(* IEC 61131-3 sources: llm-plc-st-eval/data/processed_definitivo/gpt-4o-2024-08-06/I8/zero_shot, 3 files *)

(* ---- ejec_1.st ---- *)
FUNCTION_BLOCK FB_Compresor
VAR_INPUT
    pOilOk : BOOL;        // Presión de aceite correcta
    tempOk : BOOL;        // Temperatura correcta
    sinAlm : BOOL;        // Sin alarmas
    btnMarcha : BOOL;     // Botón de marcha
    btnParo : BOOL;       // Botón de paro
END_VAR

VAR_OUTPUT
    comp : BOOL;          // Salida del compresor
    causaBloqueo : INT;   // Causa del bloqueo
END_VAR

VAR
    pOilOkTimer : TON;    // Temporizador para presión de aceite
    btnMarchaPrev : BOOL; // Estado previo del botón de marcha
END_VAR

// Inicialización del temporizador
pOilOkTimer(IN := pOilOk, PT := T#3S);

// Evaluación de los permisivos
IF NOT pOilOkTimer.Q THEN
    causaBloqueo := 1; // Falta presión de aceite
ELSIF NOT tempOk THEN
    causaBloqueo := 2; // Falta temperatura correcta
ELSIF NOT sinAlm THEN
    causaBloqueo := 3; // Alarma activa
ELSE
    causaBloqueo := 0; // Todos los permisivos están bien
END_IF

// Lógica de control del compresor
IF btnParo THEN
    comp := FALSE; // Parar el compresor
ELSIF NOT comp THEN
    // Arrancar el compresor solo si se presiona btnMarcha y todos los permisivos están bien
    IF btnMarcha AND NOT btnMarchaPrev AND causaBloqueo = 0 THEN
        comp := TRUE;
    END_IF
END_IF

// Actualizar el estado previo del botón de marcha
btnMarchaPrev := btnMarcha;
END_FUNCTION_BLOCK

(* ---- ejec_2.st ---- *)
FUNCTION_BLOCK FB_Compresor
VAR_INPUT
    pOilOk : BOOL;       // Presión de aceite correcta
    tempOk : BOOL;       // Temperatura correcta
    sinAlm : BOOL;       // Ausencia de alarmas
    btnMarcha : BOOL;    // Botón de marcha
    btnParo : BOOL;      // Botón de paro
END_VAR

VAR_OUTPUT
    comp : BOOL;         // Estado del compresor
    causaBloqueo : INT;  // Causa de bloqueo
END_VAR

VAR
    pOilOkTimer : TON;   // Temporizador para presión de aceite
    marchaPrev : BOOL;   // Estado anterior de btnMarcha
END_VAR

// Inicialización del temporizador
pOilOkTimer(IN := pOilOk, PT := T#3S);

// Lógica para determinar la causa de bloqueo
IF NOT pOilOk THEN
    causaBloqueo := 1; // Falta presión de aceite
ELSIF NOT tempOk THEN
    causaBloqueo := 2; // Falta temperatura correcta
ELSIF NOT sinAlm THEN
    causaBloqueo := 3; // Hay alarmas activas
ELSE
    causaBloqueo := 0; // No hay bloqueos
END_IF;

// Lógica de control del compresor
IF btnParo THEN
    comp := FALSE; // Parar el compresor si se pulsa btnParo
ELSIF comp THEN
    // Mantener el compresor en marcha si está en marcha y no hay bloqueos
    IF NOT (pOilOkTimer.Q AND tempOk AND sinAlm) THEN
        comp := FALSE; // Parar si se pierde algún permisivo
    END_IF;
ELSE
    // Arrancar el compresor si se pulsa btnMarcha y se cumplen los permisivos
    IF btnMarcha AND NOT marchaPrev AND pOilOkTimer.Q AND tempOk AND sinAlm THEN
        comp := TRUE;
    END_IF;
END_IF;

// Actualizar el estado anterior de btnMarcha
marchaPrev := btnMarcha;

END_FUNCTION_BLOCK

(* ---- ejec_3.st ---- *)
FUNCTION_BLOCK FB_Compresor
VAR
    // Entradas
    pOilOk : BOOL;       // Presión de aceite correcta
    tempOk : BOOL;       // Temperatura correcta
    sinAlm : BOOL;       // Sin alarmas
    btnMarcha : BOOL;    // Botón de marcha
    btnParo : BOOL;      // Botón de paro

    // Salidas
    comp : BOOL;         // Estado del compresor
    causaBloqueo : INT;  // Causa de bloqueo

    // Variables internas
    pOilOkTimer : TON;   // Temporizador para presión de aceite
    marchaLatch : BOOL;  // Latch para mantener el compresor en marcha
END_VAR

// Inicialización del temporizador
pOilOkTimer(IN := pOilOk, PT := T#3S);

// Lógica de causa de bloqueo
IF NOT pOilOkTimer.Q THEN
    causaBloqueo := 1; // Falta presión de aceite
ELSIF NOT tempOk THEN
    causaBloqueo := 2; // Falta temperatura correcta
ELSIF NOT sinAlm THEN
    causaBloqueo := 3; // Hay alarmas activas
ELSE
    causaBloqueo := 0; // No hay bloqueos
END_IF;

// Lógica de arranque y paro del compresor
IF btnParo THEN
    marchaLatch := FALSE; // Parar el compresor
ELSIF btnMarcha AND NOT marchaLatch AND (causaBloqueo = 0) THEN
    marchaLatch := TRUE; // Arrancar el compresor
END_IF;

// Actualizar el estado del compresor
comp := marchaLatch AND (causaBloqueo = 0);
